TYPE ST_WeldingPhases :
STRUCT
	stPreHeat							:ST_PreHeat;
	stBeadUp							:ST_BeadUp;
	stHeatUp							:ST_HeatUp;
	unChangeoverTime					:UINT;											(* Changeover time [s] *)
	stWelding							:ST_ForceProcess;
END_STRUCT
END_TYPE

(* stored: Version 1.1.0.1, ProductVersion 3.1.4024.15
   DUT ST_WeldingPhases: Id {066ad65c-c551-4e29-94b8-1f1873f2d7e7} *)
